// TIA Portal V21 export
VAR_GLOBAL   // PLC tag table "IO_vertikale Achse"
   ModePos_v AT %MW2 : Int;   //    {ExternalAccessible false}
   AxisEnabled_v AT %M4.4 : Bool;
   AxisPosOK_v AT %M4.0 : Bool;
   AxisRef_v AT %M4.1 : Bool;
   AxisError_v AT %M4.2 : Bool;
   Error_v AT %M4.3 : Bool;
   ActVel_v AT %M5.0 : LReal;
   ActPos_v AT %M14.0 : LReal;
END_VAR
